# EPICS substitutions: db/Beckhoff_7XXX/ecmcEX72XX_OPT_info2Inputs.substitutions
file "ecmcEL7221-9014_STD_INPUTS.template"
{
  pattern {CH_ID}
          {"$(OPT_CH_ID=01)"}
}
